FUNCTION_BLOCK FB_SignalWatchdog2
VAR_INPUT
	bEnable					:BOOL;			(* Enable FB signal *)
	bIn						:BOOL;			(* Input *)
	tTimeOutHigh				:TIME := t#5s;		(* Input high timeout *)
	tTimeOutLow				:TIME := t#5s;		(* Input low timeout *)
END_VAR
VAR_OUTPUT
	bOut					:BOOL;			(* Output *)
	bError					:BOOL;			(* Error *)
	udnErrorNo				:UDINT;
	udnMessageNo			:UDINT;
	sMsg					:STRING;
END_VAR
VAR
	bFirstTime				:BOOL;			(* First cycle *)
	tonDelay					:TON;			(* Delay *)
	tofWatchDog				:TOF;			(* Timer to off *)

END_VAR


IF NOT bFirstTime
THEN
	bError := FALSE;
	udnErrorNo := 0;
	udnMessageNo := 0;
	sMsg := '';
	tonDelay(
		IN := FALSE,
	          PT := tTimeOutHigh
	);
	tofWatchDog(
		IN := FALSE,
	         PT := tTimeOutLow
	);
	bFirstTime := TRUE;
END_IF;

(* Timer starts when came rising edge of signal *)
tonDelay(
	IN := bIn,
         PT := tTimeOutHigh
);

tofWatchDog(
	IN := bIn,
         PT := tTimeOutLow
);

IF tonDelay.Q
THEN
	bOut := TRUE;
    
ELSIF NOT tofWatchDog.Q
THEN
	bOut := FALSE;
    
END_IF;

END_FUNCTION_BLOCK

(* stored: Version 1.1.0.1, ProductVersion 3.1.4024.15
   POU FB_SignalWatchdog2: Id {9c5e3d74-c650-4048-8a47-34a4b7c05570}, SpecialFunc None *)
